SUBAPPLICATION AX_TO_Checkbox (* Gegenstueck zu Checkbox_IDA_TO_AX: AX (Pegel) auf eine VT-Checkbox schreiben (AX_TO_AD + F_DWORD_TO_UDINT + isobus::UT::Q::Q_NumericValue), schreibt bei jeder Wertaenderung von AX_IN neu auf den VT-Knoten. WICHTIG: u16ObjId ist die ObjectID der CNumberVariable, die die Checkbox als Wertspeicher referenziert (z.B. NumberVariable_Bunker_Fuellstand_Hoehe_Automatik) - NICHT die ObjectID der Checkbox (CInputBoolean) selbst, die VT erwartet Value-Aenderungen unter der NumberVariable-ID (analog Checkbox_IDA_TO_AX, Franz, live verifiziert). Instanz-Eindeutigkeit beachten: Q_NumericValue erlaubt nur eine Instanz je Ziel-ObjId im gesamten Projekt. *)
  (* Standard: 61499-2; Description: Copyright (c) 2026 Büngener Schuder GmbH This program and the accompanying materials are made available under the terms of the Eclipse Public License 2.0 which is available at https://www.eclipse.org/legal/epl-2.0/ SPDX-License-Identifier: EPL-2.0 *)
  (* Version 1.0, 2026-10-13, Franz Höpfinger, Büngener Schuder GmbH, initial implementation - Gegenstelle zu Checkbox_IDA_TO_AX (ECU->VT statt VT->ECU). AX_TO_AD (bit-reinterpretiert BOOL->DWORD, feuert nur bei echter Wertaenderung) -> F_DWORD_TO_UDINT -> Q_NumericValue.REQ, analog zu Q_NumericValue_AUDI's eigenem u32NewValue-Adapter-Socket-Muster (isobus_UT_adapter), nur ohne eigenen Adapter-Typ dafuer - hier als SubApp-Komposition. *)
  PACKAGE MyLib::sys;
  IMPORT isobus::UT::Q::const::IDs::ID_NULL;
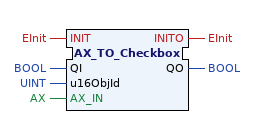
  EVENT_INPUT
    INIT : EInit; (* Initialization Request *)
  END_EVENT
  EVENT_OUTPUT
    INITO : EInit; (* Initialization Confirm *)
  END_EVENT
  VAR_INPUT
    QI : BOOL := TRUE; (* Quality Input - TRUE to enable service *)
    u16ObjId : UINT := ID_NULL; (* Object ID der VT-NumberVariable hinter der Checkbox *)
  END_VAR
  VAR_OUTPUT
    QO : BOOL; (* Quality Output - TRUE if service executed successfully *)
  END_VAR
  SOCKETS
    AX_IN : adapter::types::unidirectional::AX; (* Zu schreibender Pegel (0/1) *)
  END_SOCKETS
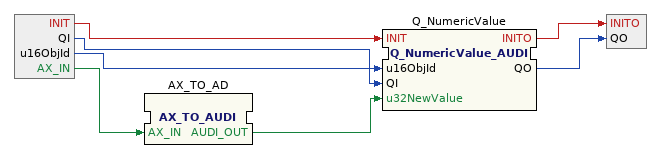
  FBS
    AX_TO_AD : adapter::conversion::unidirectional::AX_TO_AUDI;
    Q_NumericValue : isobus::UT::Q::Q_NumericValue_AUDI;
  END_FBS
  EVENT_CONNECTIONS
    INIT TO Q_NumericValue.INIT;
    Q_NumericValue.INITO TO INITO;
  END_CONNECTIONS
  DATA_CONNECTIONS
    u16ObjId TO Q_NumericValue.u16ObjId;
    QI TO Q_NumericValue.QI;
    Q_NumericValue.QO TO QO;
  END_CONNECTIONS
  ADAPTER_CONNECTIONS
    AX_IN TO AX_TO_AD.AX_IN;
    AX_TO_AD.AUDI_OUT TO Q_NumericValue.u32NewValue;
  END_CONNECTIONS
END_SUBAPPLICATION
